// TIA Portal V20 export
FUNCTION_BLOCK "FB_Valve"   // FB101, LAD
TITLE = On/off valve with limit switch monitoring
{ S7_Optimized_Access := 'TRUE' }
AUTHOR : Demo
VERSION : 0.2
// LAD version. Same interface as scl/13_FB_Valve.scl.
// stored: AutoNumber false, SetENOAutomatically false
   VAR_INPUT
      Open : Bool;   // Request: open the valve
      Permit : Bool := true;   // Interlock: valve may only open when TRUE
      ZSO : Bool;   // Open limit switch
      ZSC : Bool;   // Closed limit switch
      MonitorTime : Time := T#10S;   // Max travel time before a fault
   END_VAR
   VAR_OUTPUT
      Out : Bool;   // Open command to the solenoid
      IsOpen : Bool;   // Valve confirmed open
      IsClosed : Bool;   // Valve confirmed closed
      FaultNotOpen : Bool;   // Open command on, but open limit switch not reached in MonitorTime
      FaultNotClosed : Bool;   // Open command off, but closed limit switch not reached in MonitorTime
   END_VAR
   VAR
      tOpen : TON_TIME;   // Opening travel time
      tClose : TON_TIME;   // Closing travel time
   END_VAR
BEGIN

REGION Network 1: Open command
   // The solenoid gets the open command only when the sequence asks for it and the interlock permits it.
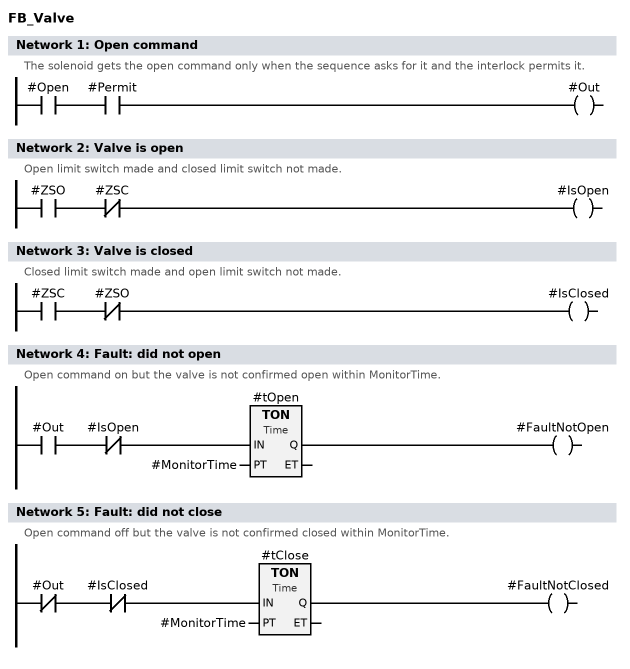
   RUNG wire#powerrail
      Contact( #Open )
      Contact( #Permit )
      Coil( #Out )
   END_RUNG
   // the same network as SCL:
   #Out := #Open AND #Permit;
END_REGION

REGION Network 2: Valve is open
   // Open limit switch made and closed limit switch not made.
   RUNG wire#powerrail
      Contact( #ZSO )
      I_Contact( #ZSC )
      Coil( #IsOpen )
   END_RUNG
   // the same network as SCL:
   #IsOpen := #ZSO AND NOT #ZSC;
END_REGION

REGION Network 3: Valve is closed
   // Closed limit switch made and open limit switch not made.
   RUNG wire#powerrail
      Contact( #ZSC )
      I_Contact( #ZSO )
      Coil( #IsClosed )
   END_RUNG
   // the same network as SCL:
   #IsClosed := #ZSC AND NOT #ZSO;
END_REGION

REGION Network 4: Fault: did not open
   // Open command on but the valve is not confirmed open within MonitorTime.
   RUNG wire#powerrail
      Contact( #Out )
      I_Contact( #IsOpen )
      { S7_Templates := "time_type := Time" } #tOpen.TON(pt := #MonitorTime, et =>)
      Coil( #FaultNotOpen )
   END_RUNG
   // the same network as SCL:
   #tOpen(IN := #Out AND NOT #IsOpen, PT := #MonitorTime);   // TON
   #FaultNotOpen := #tOpen.Q;
END_REGION

REGION Network 5: Fault: did not close
   // Open command off but the valve is not confirmed closed within MonitorTime.
   RUNG wire#powerrail
      I_Contact( #Out )
      I_Contact( #IsClosed )
      { S7_Templates := "time_type := Time" } #tClose.TON(pt := #MonitorTime, et =>)
      Coil( #FaultNotClosed )
   END_RUNG
   // the same network as SCL:
   #tClose(IN := NOT #Out AND NOT #IsClosed, PT := #MonitorTime);   // TON
   #FaultNotClosed := #tClose.Q;
END_REGION
END_FUNCTION_BLOCK
